TYPE ST_AxisParameter :
STRUCT
	/// Axis ID 
	nAxisId: DWORD;
	fLength: LREAL;
	fClampLength: LREAL;
	fGap: LREAL;
	stRoadParam: ST_RoadParameter;
	stDynamicDefault: ST_DynamicDefaultAxis;
END_STRUCT
END_TYPE

(* stored: Version 1.1.0.1, ProductVersion 3.1.4024.12
   DUT ST_AxisParameter: Id {8c28c0cc-89b6-4379-8c02-26ecbd590988} *)
